INTERFACE I_IoGroup EXTENDS I_IoBase

METHOD AddIo
VAR_INPUT
	bIo		: I_IoBit;
END_VAR
END_METHOD

END_INTERFACE

(* stored: Version 1.1.0.1
   Itf I_IoGroup: Id {43e5735c-166e-471f-b546-8f72f9ab0af3}
   Method AddIo: Id {7044145b-f295-45a4-b20f-5bbba23c3e73} *)
